// TIA Portal V20 export
// export: Created 2026-10-20T12:45:00.9116663Z, ExportSetting WithDefaults, DisplayName Totally Integrated Automation Portal, DisplayVersion V20 Update 6, DisplayName TIA Portal Openness, DisplayVersion V20 Update 6, DisplayName TIA Portal Version Control Interface, DisplayVersion V20 Update 6, DisplayName SINAMICS Startdrive Advanced, DisplayVersion V20 SP1, DisplayName SINAMICS Startdrive G130, G150, S120, S150, SINAMICS MV, G220, S200, S210, DisplayVersion V20 SP1, DisplayName SINAMICS Startdrive G110M, G120, G120C, G120D, G120P, G115D, DisplayVersion V20 SP1, DisplayName STEP 7 Professional, DisplayVersion V20 Update 6, DisplayName STEP 7 Safety, DisplayVersion V20 Update 2, DisplayName WinCC Basic/Comfort/Advanced, DisplayVersion V20 Update 6, DisplayName WinCC Unified, DisplayVersion V20 Update 6
FUNCTION "Settings_Limits_FC" : Void   // FC65, SCL
{ S7_Optimized_Access := 'TRUE' }
VERSION : 0.1
// stored: AutoNumber true, IsIECCheckEnabled false, SetENOAutomatically false, UDAEnableTagReadback false
   VAR_IN_OUT
      VTD_Settings : "VTD_Settings";
   END_VAR
BEGIN
   IF #VTD_Settings.Lowest_Level < 1 THEN
       #VTD_Settings.Lowest_Level := 1;
   END_IF;

   IF #VTD_Settings.Highest_Level > 8 THEN
       #VTD_Settings.Lowest_Level := 8;
   END_IF;

   IF #VTD_Settings.Creep_Speed < 3 THEN
       #VTD_Settings.Creep_Speed := 3;
   END_IF;

   IF #VTD_Settings.Slow_Speed < 3 THEN
       #VTD_Settings.Slow_Speed := 3;
   END_IF;

   IF #VTD_Settings.Loaded_Speed < #VTD_Settings.Slow_Calib_Speed * 1.8 THEN
       #VTD_Settings.Loaded_Speed := #VTD_Settings.Slow_Calib_Speed * 1.8;
   END_IF;

   IF #VTD_Settings.Shuttle_Speed < #VTD_Settings.Slow_Calib_Speed * 1.8 THEN
       #VTD_Settings.Shuttle_Speed := #VTD_Settings.Slow_Calib_Speed * 1.8;
   END_IF;

   IF #VTD_Settings.Pallet_Speed < #VTD_Settings.Slow_Calib_Speed * 1.8 THEN
       #VTD_Settings.Pallet_Speed := #VTD_Settings.Slow_Calib_Speed * 1.8;
   END_IF;

   IF #VTD_Settings.Empty_Speed < #VTD_Settings.Slow_Calib_Speed * 1.8 THEN
       #VTD_Settings.Empty_Speed := #VTD_Settings.Slow_Calib_Speed * 1.8;
   END_IF;

   IF #VTD_Settings.Dock_speed > 10 THEN
       #VTD_Settings.Dock_speed := 10;
   END_IF;

   IF #VTD_Settings.Empty_Speed > 120 THEN
       #VTD_Settings.Empty_Speed := 120;
   END_IF;

   IF #VTD_Settings.Pallet_Speed > 120 THEN
       #VTD_Settings.Pallet_Speed := 120;
   END_IF;

   IF #VTD_Settings.Chain_Slack_Timeout > 5000 THEN
       #VTD_Settings.Chain_Slack_Timeout := 5000;
   END_IF;

   IF #VTD_Settings.Acc_Range_1 < 60 THEN
       #VTD_Settings.Acc_Range_1 := 60;
   END_IF;

   IF #VTD_Settings.Acc_Range_2 < 60 THEN
       #VTD_Settings.Acc_Range_2 := 60;
   END_IF;

   IF #VTD_Settings.Acc_Range_3 < 60 THEN
       #VTD_Settings.Acc_Range_3 := 60;
   END_IF;

   IF #VTD_Settings.Acc_Range_1 > 100 THEN
       #VTD_Settings.Acc_Range_1 := 100;
   END_IF;

   IF #VTD_Settings.Acc_Range_2 > 100 THEN
       #VTD_Settings.Acc_Range_2 := 100;
   END_IF;

   IF #VTD_Settings.Acc_Range_3 > 100 THEN
       #VTD_Settings.Acc_Range_3 := 100;
   END_IF;
END_FUNCTION
